// TIA Portal V20 export
Screen "OP03Pop-up_PRBWork"  274x181
  ScreenItem "Text field TG Status" at 1,0 size 273x47  Type=HmiTextBox
  ScreenItem "Cancel Mode" at 195,3 size 76x42  Type=HmiButton
  ScreenItem "Rectangle TG1" at 4,52 size 265x29  Type=HmiRectangle
  ScreenItem "Textfeld_1" at 9,57 size 21x20  Type=HmiTextBox
  ScreenItem "Textfeld_2" at 50,56 size 245x20  Type=HmiTextBox
  ScreenItem "Rectangle TG1_1" at 4,84 size 265x29  Type=HmiRectangle
  ScreenItem "Textfeld_5" at 9,88 size 21x20  Type=HmiTextBox
  ScreenItem "Rectangle TG1_2" at 4,116 size 265x29  Type=HmiRectangle
  ScreenItem "Rectangle TG1_3" at 4,148 size 265x29  Type=HmiRectangle
  ScreenItem "Textfeld_3" at 50,88 size 245x20  Type=HmiTextBox
  ScreenItem "Textfeld_16" at 9,121 size 21x20  Type=HmiTextBox
  ScreenItem "Textfeld_13" at 50,120 size 275x20  Type=HmiTextBox
  ScreenItem "Line_1" at 37,52 size 0x125  Type=HmiLine
  ScreenItem "Textfeld_4" at 9,152 size 21x20  Type=HmiTextBox
  ScreenItem "Textfeld_6" at 50,152 size 275x20  Type=HmiTextBox
